(* IEC 61131-3 sources: volt/packages/volt-lsp-iec/test-corpus/pro2193/Device/Plc Logic/Application/09 Misc/Library Manager/CommFB, 61 files *)

(* ---- ADDR_TYPE.dut ---- *)
TYPE ADDR_TYPE :
UNION
	SYSTEM : IO_SYSTEM_TYPE;
	DP : DP_ADDR;
	PN : PN_ADDR;
END_UNION
END_TYPE

(* ---- AINFO_TYPE.dut ---- *)
TYPE AINFO_TYPE :
UNION
	DP : DP_AINFO;
	PN : PN_AINFO;
END_UNION
END_TYPE

(* ---- CNCT_STATE.dut ---- *)
TYPE CNCT_STATE :
(
	S1_INIT := 1,
	S2_IDLE := 2,
	S3_CONNECTING := 3,
	S4_CONNECTED := 4,
	S5_DISCONNECTING := 5,
	S6_ERROR := 6
);
END_TYPE

(* ---- DP_ADDR.dut ---- *)
TYPE DP_ADDR :
STRUCT
	SYSTEM : IO_SYSTEM_TYPE;
	VERSION : BYTE := 1;
	D : DP_DEVICE_ID;
	SLOT : BYTE;
END_STRUCT
END_TYPE

(* ---- DP_AINFO.dut ---- *)
TYPE DP_AINFO :
STRUCT
	D_LEN : BYTE;
	ATYPE : BYTE;
	SLOT : BYTE;
	ASPEC : BYTE;
	ADD_INFO : ARRAY [0..58] OF BYTE;
END_STRUCT
END_TYPE

(* ---- DP_DEVICE_ID.dut ---- *)
TYPE DP_DEVICE_ID :
STRUCT
	MASTER : BYTE;
	SEGMENT : BYTE;
	STATION : BYTE;
END_STRUCT
END_TYPE

(* ---- DP_DIAG.dut ---- *)
TYPE DP_DIAG :
STRUCT
	STATUS1 : IIoDrvProfibus.DP_StationStatus1;
	STATUS2 : IIoDrvProfibus.DP_StationStatus2;
	STATUS3 : IIoDrvProfibus.DP_StationStatus3;
	DIAG_MASTER_ADD : USINT;
	IDENT_NUMBER : UINT;
	EXTDIAG : ARRAY [0..235] OF BYTE;
END_STRUCT
END_TYPE

(* ---- ERRORCODE.dut ---- *)
TYPE ERRORCODE :
(
	NONE := 0,
	INVALID_ID := 16#40820000,
	UNKNOWN := 16#40000100,
	NOT_IMPLEMENTED := 16#40000101,
	RDIAG_PROFINET := 16#40000102,
	STACK_NOT_RUNNING := 16#40000103,
	NO_RESSOURCE := 16#40000104,
	BUFFER_SIZE := 16#40000105,
	INVALID_STATE := 16#40000110,
	ADDRESS_NOT_UNIQUE := 16#40000111,
	ADDRESS_INVALID := 16#40000112,
	DEVICE_NOT_FOUND := 16#40000113,
	DEVICETYPE_MISMATCH := 16#40000114,
	TIMEOUT := 16#40000115
);
END_TYPE

(* ---- ERRORCODE1_RW.dut ---- *)
TYPE ERRORCODE1_RW :
(
	INVALID_INDEX := 16#B0,
	WRITE_LENGTH_ERROR := 16#B1,
	INVALID_SLOT_OR_SUBSLOT := 16#B2,
	TYPE_CONFLICT := 16#B3,
	INVALID_AREA_OR_API := 16#B4,
	STATE_CONFLICT := 16#B5,
	ACCESS_DENIED := 16#B6,
	INVALID_RANGE := 16#B7,
	INVALID_PARAMETER := 16#B8,
	INVALID_TYPE := 16#B9,
	BACKUP := 16#BA
);
END_TYPE

(* ---- IO_SYSTEM_TYPE.dut ---- *)
TYPE IO_SYSTEM_TYPE :
(
	PROFIBUS_DP := 1,
	PROFINET_IO := 2
);
END_TYPE

(* ---- PN_ADDR.dut ---- *)
TYPE PN_ADDR :
STRUCT
	SYSTEM : IO_SYSTEM_TYPE;
	VERSION : BYTE := 1;
	MASTER : BYTE;
	D : PN_DEVICE_ID;
	API : DWORD;
	SLOT : WORD;
	SUBSLOT : WORD;
END_STRUCT
END_TYPE

(* ---- PN_AINFO.dut ---- *)
TYPE PN_AINFO :
STRUCT
	BLOCKTYPE : UINT;
	BLOCKLENGTH : UINT;
	VERSION : UINT;
	ALARMTYPE : UINT;
	API : UDINT;
	SLOT : UINT;
	SUBSLOT : UINT;
	MODULEIDENTNUMBER : UDINT;
	SUBMODULEIDENTNUMBER : UDINT;
	ALARMSPECIFIER : UINT;
	USI : UINT;
	ALARMDATA : ARRAY [0..(Constants.MAX_PN_ALARM_DATA - 1)] OF BYTE;
END_STRUCT
END_TYPE

(* ---- PN_DEVICE_ID.dut ---- *)
TYPE PN_DEVICE_ID :
STRUCT
	STATIONNAME : STRING;
	INSTANCE : WORD;
	DEVICE : WORD;
	VENDOR : WORD;
END_STRUCT
END_TYPE

(* ---- PRVREC_MODE.dut ---- *)
TYPE PRVREC_MODE :
(
	CHECK := 0,
	RECEIVE := 1,
	RECEIVE_BY_SLOT := 2,
	POS_RESPONSE := 3,
	NEG_RESPONSE := 4
);
END_TYPE

(* ---- PRVREC_STATE.dut ---- *)
TYPE PRVREC_STATE :
(
	S1_INIT,
	S2_IDLE,
	S3_ENABLED,
	S4_NEG_RESP,
	S5_RECEIVED,
	S6_CHECK,
	S7_POS_RESP,
	S8_NEG_RESP,
	S9_ERROR
);
END_TYPE

(* ---- RALARM_MODE.dut ---- *)
TYPE RALARM_MODE :
(
	ALL_ALARMS := 1,
	ALARM_BY_ID := 2,
	ALARM_BY_SLOT := 3,
	ALARM_BY_DEVICE := 4
);
END_TYPE

(* ---- RCVREC_MODE.dut ---- *)
TYPE RCVREC_MODE :
(
	CHECK := 0,
	RECEIVE := 1,
	RECEIVE_BY_SLOT := 2,
	POS_RESPONSE := 3,
	NEG_RESPONSE := 4
);
END_TYPE

(* ---- RCVREC_STATE.dut ---- *)
TYPE RCVREC_STATE :
(
	S1_INIT,
	S2_IDLE,
	S3_ENABLED,
	S4_NEG_RESP,
	S5_RECEIVED,
	S6_CHECK,
	S7_POS_RESP,
	S8_NEG_RESP,
	S9_ERROR
);
END_TYPE

(* ---- RDREC_STATE.dut ---- *)
TYPE RDREC_STATE :
(
	S1_INIT := 1,
	S2_IDLE := 2,
	S3_WAITING := 3,
	S4_HAVEDATA := 4,
	S5_ERROR := 5
);
END_TYPE

(* ---- READ_IND.dut ---- *)
TYPE READ_IND :
STRUCT
	SLOT : UINT;
	SUBSLOT : UINT;
	INDEX : UINT;
	RLEN : UINT;
	AR_ID : DWORD;
	SEQ_NUMBER : UINT;
END_STRUCT
END_TYPE

(* ---- SALRM_STATE.dut ---- *)
TYPE SALRM_STATE :
(
	S1_INIT,
	S2_IDLE,
	S3_WAITING,
	S4_HAVE_ACK,
	S5_ERROR
);
END_TYPE

(* ---- WRITE_IND.dut ---- *)
TYPE WRITE_IND :
STRUCT
	SLOT : UINT;
	SUBSLOT : UINT;
	INDEX : UINT;
	PRM : BOOL;
	AR_ID : DWORD;
	SEQ_NUMBER : UINT;
	LEN : UINT;
	DATA : POINTER TO BYTE;
END_STRUCT
END_TYPE

(* ---- WRREC_STATE.dut ---- *)
TYPE WRREC_STATE :
(
	S1_INIT := 1,
	S2_IDLE := 2,
	S3_WAITING := 3,
	S4_DATAWRITTEN := 4,
	S5_ERROR := 5
);
END_TYPE

(* ---- ADDRESSCONCEPT.gvl ---- *)
VAR_GLOBAL
	DUMMY : UDINT := 0;
END_VAR

(* ---- CONSTANTS.gvl ---- *)
VAR_GLOBAL
	INVALID_ID : UDINT := 16#FFFFFFFF;
	MAX_PN_ALARM_DATA : UDINT := 198;
END_VAR

(* ---- ICOMMFBALARMSENDER.itf ---- *)
INTERFACE ICOMMFBALARMSENDER
END_INTERFACE

METHOD ALARMCNF
VAR_INPUT
	ERROR : DWORD;
END_VAR
END_METHOD

(* ---- ICOMMFBCONNECTIONMANAGERFACTORY.itf ---- *)
INTERFACE ICOMMFBCONNECTIONMANAGERFACTORY
END_INTERFACE

METHOD GETCONNECTIONMANAGER : UDINT
VAR_INPUT
	CLIENT : IConnectionManagerClient;
END_VAR
VAR_OUTPUT
	CONNECTIONMANAGER : IConnectionManager;
END_VAR
VAR_IN_OUT
	D_ADDR : ADDR_TYPE;
END_VAR
END_METHOD

METHOD RELEASECONNECTIONMANAGER : UDINT
VAR_INPUT
	CLIENT : IConnectionManagerClient;
	CONNECTIONMANAGER : IConnectionManager;
END_VAR
END_METHOD

(* ---- ICOMMFBDIAGPROVIDER.itf ---- *)
INTERFACE ICOMMFBDIAGPROVIDER
END_INTERFACE

METHOD CHECKOWNER : BOOL
VAR_INPUT
	ID : UDINT;
END_VAR
END_METHOD

METHOD GETALARM : DWORD
VAR_INPUT
	MODE : INT;
	F_ID : DWORD;
END_VAR
VAR_OUTPUT
	NEW : BOOL;
	ID : DWORD;
	LEN : INT;
END_VAR
VAR_IN_OUT
	AINFO : AINFO_TYPE;
	CURRENTALARMID : UDINT;
END_VAR
END_METHOD

METHOD GETDIAG : DWORD
VAR_INPUT
	ID : DWORD;
END_VAR
VAR_OUTPUT
	BUSY : BOOL;
	LEN : INT;
END_VAR
VAR_IN_OUT
	DINFO : DP_DIAG;
END_VAR
END_METHOD

(* ---- ICOMMFBFACTORY.itf ---- *)
INTERFACE ICOMMFBFACTORY
END_INTERFACE

METHOD CHECKOWNER : BOOL
VAR_INPUT
	ID : UDINT;
END_VAR
END_METHOD

METHOD GETRDREC : POINTER TO RDRECBase
VAR_INPUT
	ID : UDINT;
END_VAR
VAR_IN_OUT
	CLIENT : RDREC;
END_VAR
END_METHOD

METHOD GETWRREC : POINTER TO WRRECBase
VAR_INPUT
	ID : UDINT;
END_VAR
VAR_IN_OUT
	CLIENT : WRREC;
END_VAR
END_METHOD

METHOD RELEASERDREC : BOOL
VAR_INPUT
	ID : UDINT;
END_VAR
VAR_IN_OUT
	CLIENT : RDREC;
END_VAR
END_METHOD

METHOD RELEASEWRREC : BOOL
VAR_INPUT
	ID : UDINT;
END_VAR
VAR_IN_OUT
	CLIENT : WRREC;
END_VAR
END_METHOD

(* ---- ICOMMFBFACTORYEXT.itf ---- *)
INTERFACE ICOMMFBFACTORYEXT
END_INTERFACE

METHOD TRYGETADDRESS : BOOL
VAR_INPUT
	ID : DWORD;
END_VAR
VAR_OUTPUT
	STATUS : DWORD;
END_VAR
VAR_IN_OUT
	ADDR : ADDR_TYPE;
END_VAR
END_METHOD

METHOD TRYGETID : BOOL
VAR_OUTPUT
	STATUS : DWORD;
	ID : DWORD;
END_VAR
VAR_IN_OUT
	ADDR : ADDR_TYPE;
END_VAR
END_METHOD

(* ---- ICOMMFBFACTORYIO.itf ---- *)
INTERFACE ICOMMFBFACTORYIO
END_INTERFACE

METHOD CHECKOWNER : BOOL
VAR_INPUT
	ID : UDINT;
END_VAR
END_METHOD

METHOD GETINPUTDATA : DWORD
VAR_INPUT
	ID : DWORD;
	OFFSET : UINT;
	LEN : UINT;
	INPUTS : POINTER TO BYTE;
END_VAR
VAR_OUTPUT
	IO_LEN : UINT;
	CONSISTENCY : BOOL;
END_VAR
END_METHOD

METHOD PUTOUTPUTDATA : DWORD
VAR_INPUT
	ID : DWORD;
	OFFSET : UINT;
	LEN : UINT;
	OUTPUTS : POINTER TO BYTE;
END_VAR
VAR_OUTPUT
	IO_LEN : UINT;
	CONSISTENCY : BOOL;
END_VAR
END_METHOD

(* ---- ICOMMFBFIELDDEVICE.itf ---- *)
INTERFACE ICOMMFBFIELDDEVICE
END_INTERFACE

METHOD ALARMREQ : DWORD
VAR_INPUT
	ALARMSENDER : ICommFBAlarmSender;
	ID : DWORD;
	ATYPE : UINT;
	ASPEC : UINT;
	LEN : UINT;
	AINFO : POINTER TO BYTE;
END_VAR
END_METHOD

METHOD CHECKREADIND : BOOL
VAR_INPUT
	MODE : UINT;
	F_ID : DWORD;
END_VAR
VAR_OUTPUT
	STATUS : DWORD;
	IND : Read_Ind;
END_VAR
END_METHOD

METHOD CHECKWRITEIND : BOOL
VAR_INPUT
	MODE : UINT;
	F_ID : DWORD;
END_VAR
VAR_OUTPUT
	STATUS : DWORD;
	IND : Write_Ind;
END_VAR
END_METHOD

METHOD READNEGRSP : DWORD
VAR_INPUT
	CODE1 : BYTE;
	CODE2 : BYTE;
END_VAR
VAR_IN_OUT
	IND : Read_Ind;
END_VAR
END_METHOD

METHOD READRSP : DWORD
VAR_INPUT
	LEN : UINT;
	RECORD : POINTER TO BYTE;
END_VAR
VAR_IN_OUT
	IND : Read_Ind;
END_VAR
END_METHOD

METHOD WRITENEGRSP : DWORD
VAR_INPUT
	CODE1 : BYTE;
	CODE2 : BYTE;
END_VAR
VAR_IN_OUT
	IND : Write_Ind;
END_VAR
END_METHOD

METHOD WRITERSP : DWORD
VAR_IN_OUT
	IND : Write_Ind;
END_VAR
END_METHOD

(* ---- ICONNECTIONMANAGER.itf ---- *)
INTERFACE ICONNECTIONMANAGER
END_INTERFACE

METHOD CONNECTREQ : DWORD
VAR_IN_OUT
	D_ADDR : ADDR_TYPE;
END_VAR
END_METHOD

METHOD RELEASEREQ : DWORD
END_METHOD

METHOD UPDATEADDRESS : DWORD
VAR_IN_OUT
	D_ADDR : ADDR_TYPE;
END_VAR
END_METHOD

(* ---- ICONNECTIONMANAGERCLIENT.itf ---- *)
INTERFACE ICONNECTIONMANAGERCLIENT
END_INTERFACE

METHOD CONNECTCNF
VAR_INPUT
	ID : DWORD;
	ERRORCODE : DWORD;
END_VAR
END_METHOD

METHOD ERRORIND
VAR_INPUT
	ERRORCODE : DWORD;
END_VAR
END_METHOD

METHOD RELEASECNF
VAR_INPUT
	ERRORCODE : DWORD;
END_VAR
END_METHOD

(* ---- IGENERICIDFACTORY.itf ---- *)
INTERFACE IGENERICIDFACTORY
END_INTERFACE

METHOD TRYGETIDFROMREFERENCE : BOOL
VAR_INPUT
	PREF : POINTER TO BYTE;
END_VAR
VAR_OUTPUT
	ID : DWORD;
END_VAR
END_METHOD

(* ---- ADDR.pou ---- *)
FUNCTION ADDR : DWORD
VAR_INPUT
	EN : BOOL := TRUE;
	ID : DWORD;
END_VAR
VAR_OUTPUT
	ENO : BOOL;
END_VAR
END_FUNCTION

(* ---- ID.pou ---- *)
FUNCTION ID : DWORD
VAR_INPUT
	EN : BOOL := TRUE;
	MASTER : BYTE;
	SEGMENT : BYTE;
	STATION : BYTE;
	SLOT : BYTE;
END_VAR
END_FUNCTION

(* ---- ID_FROM_REF.pou ---- *)
FUNCTION ID_FROM_REF : DWORD
VAR_INPUT
	PREF : POINTER TO BYTE;
END_VAR
END_FUNCTION

(* ---- SLOT_ID.pou ---- *)
FUNCTION SLOT_ID : DWORD
VAR_INPUT
	EN : BOOL := TRUE;
	ID : DWORD;
	SLOT : BYTE;
END_VAR
VAR_OUTPUT
	ENO : BOOL;
END_VAR
END_FUNCTION

(* ---- SUBSLOT_ID.pou ---- *)
FUNCTION SUBSLOT_ID : DWORD
VAR_INPUT
	EN : BOOL := TRUE;
	ID : DWORD;
	SLOT : UINT;
	SUBSLOT : UINT;
END_VAR
VAR_OUTPUT
	ENO : BOOL;
END_VAR
END_FUNCTION

(* ---- ADDR_TO_ID.pou ---- *)
FUNCTION_BLOCK ADDR_TO_ID
VAR_INPUT
	EN : BOOL := TRUE;
END_VAR
VAR_OUTPUT
	ENO : BOOL;
	STATUS : DWORD;
	ID : DWORD;
END_VAR
VAR_IN_OUT
	ADDR : ADDR_TYPE;
END_VAR
VAR
	S_INSTANCEHANDLER : InstanceHandler;
	I : DINT;
END_VAR
END_FUNCTION_BLOCK

(* ---- ALARMSENDERINTERNAL.pou ---- *)
FUNCTION_BLOCK ALARMSENDERINTERNAL
VAR_INPUT
	SALARM : POINTER TO SALARM;
END_VAR
END_FUNCTION_BLOCK

METHOD ALARMCNF
VAR_INPUT
	ERROR : DWORD;
END_VAR
END_METHOD

(* ---- CNCT.pou ---- *)
FUNCTION_BLOCK CNCT
VAR_INPUT
	REQ : BOOL;
	D_ADDR : ADDR_TYPE;
END_VAR
VAR_OUTPUT
	VALID : BOOL;
	ERROR : BOOL;
	BUSY : BOOL;
	STATUS : DWORD;
	ID : DWORD := Constants.INVALID_ID;
END_VAR
VAR
	S_INSTANCEHANDLER : InstanceHandler;
	_FACTORY : ICommFBConnectionManagerFactory;
	_CONNECTIONMANAGER : IConnectionManager;
	_REQ : BOOL;
	_STATE : CNCT_State := CNCT_State.S2_Idle;
	_ERRORCODE : UDINT;
	_CONNECTREQ : UDINT;
	_CONNECTID : DWORD := Constants.INVALID_ID;
	_RECVCONNECTCNF : BOOL;
	_RECVRELEASECNF : BOOL;
	_RECVABORTIND : BOOL;
	_CLIENT : ConnectionManagerClientInternal;
END_VAR
END_FUNCTION_BLOCK

METHOD ABORTIND
VAR_INPUT
	ERRORCODE : DWORD;
END_VAR
END_METHOD

METHOD CONNECTCNF
VAR_INPUT
	ID : DWORD;
	ERRORCODE : DWORD;
END_VAR
END_METHOD

METHOD RELEASECNF
VAR_INPUT
	ERRORCODE : DWORD;
END_VAR
END_METHOD

(* ---- CONNECTIONMANAGERCLIENTIMPLICITID.pou ---- *)
FUNCTION_BLOCK CONNECTIONMANAGERCLIENTIMPLICITID
VAR_INPUT
	CNCT : POINTER TO CREATE_ID;
END_VAR
END_FUNCTION_BLOCK

METHOD CONNECTCNF
VAR_INPUT
	ID : DWORD;
	ERRORCODE : DWORD;
END_VAR
END_METHOD

METHOD ERRORIND
VAR_INPUT
	ERRORCODE : DWORD;
END_VAR
END_METHOD

METHOD RELEASECNF
VAR_INPUT
	ERRORCODE : DWORD;
END_VAR
END_METHOD

(* ---- CONNECTIONMANAGERCLIENTINTERNAL.pou ---- *)
FUNCTION_BLOCK CONNECTIONMANAGERCLIENTINTERNAL
VAR_INPUT
	CNCT : POINTER TO CNCT;
END_VAR
END_FUNCTION_BLOCK

METHOD CONNECTCNF
VAR_INPUT
	ID : DWORD;
	ERRORCODE : DWORD;
END_VAR
END_METHOD

METHOD ERRORIND
VAR_INPUT
	ERRORCODE : DWORD;
END_VAR
END_METHOD

METHOD RELEASECNF
VAR_INPUT
	ERRORCODE : DWORD;
END_VAR
END_METHOD

(* ---- CREATE_ID.pou ---- *)
FUNCTION_BLOCK CREATE_ID
VAR_INPUT
	EN : BOOL := TRUE;
END_VAR
VAR_OUTPUT
	ENO : BOOL;
	STATUS : DWORD;
	ID : DWORD;
END_VAR
VAR_IN_OUT
	ADDR : ADDR_TYPE;
END_VAR
VAR
	S_INSTANCEHANDLER : InstanceHandler;
	_FACTORY : ICommFBConnectionManagerFactory;
	_CONNECTIONMANAGER : IConnectionManager;
	_STATE : CNCT_State := CNCT_State.S2_Idle;
	_ERRORCODE : UDINT;
	_CONNECTID : DWORD := Constants.INVALID_ID;
	_RECVCONNECTCNF : BOOL;
	_RECVRELEASECNF : BOOL;
	_RECVABORTIND : BOOL;
	_CLIENT : ConnectionManagerClientImplicitID;
	D_ADDR : ADDR_TYPE;
END_VAR
END_FUNCTION_BLOCK

METHOD ABORTIND
VAR_INPUT
	ERRORCODE : DWORD;
END_VAR
END_METHOD

METHOD CONNECTCNF
VAR_INPUT
	ID : DWORD;
	ERRORCODE : DWORD;
END_VAR
END_METHOD

METHOD RELEASECNF
VAR_INPUT
	ERRORCODE : DWORD;
END_VAR
END_METHOD

(* ---- GETIO_PART.pou ---- *)
FUNCTION_BLOCK GETIO_PART
VAR_INPUT
	EN : BOOL;
	ID : DWORD;
	OFFSET : INT;
	LEN : INT;
	INPUTS : POINTER TO BYTE;
END_VAR
VAR_OUTPUT
	ENO : BOOL;
	STATUS : DWORD;
	ERROR : BOOL;
END_VAR
VAR
	S_INSTANCEHANDLER : InstanceHandler;
	I : DINT;
	_FACTORY : ICommFBFactoryIO;
	IOLEN : UINT;
	TRANSFERCONSISTENT : BOOL;
END_VAR
END_FUNCTION_BLOCK

(* ---- ID_TO_ADDR.pou ---- *)
FUNCTION_BLOCK ID_TO_ADDR
VAR_INPUT
	EN : BOOL := TRUE;
	ID : DWORD;
END_VAR
VAR_OUTPUT
	ENO : BOOL;
	STATUS : DWORD;
END_VAR
VAR_IN_OUT
	ADDR : ADDR_TYPE;
END_VAR
VAR
	S_INSTANCEHANDLER : InstanceHandler;
	I : DINT;
	FACTORY : ICommFBFactoryExt;
END_VAR
END_FUNCTION_BLOCK

(* ---- INSTANCEHANDLER.pou ---- *)
FUNCTION_BLOCK INSTANCEHANDLER
VAR
	S_INSTANCECOUNT : UINT;
	S_FACTORIES : ARRAY [0..(MAX_INSTANCES - 1)] OF ICommFBFactory;
	S_FACTORIESEXT : ARRAY [0..(MAX_INSTANCES - 1)] OF ICommFBFactoryExt;
	S_FACTORIESIO : ARRAY [0..(MAX_INSTANCES - 1)] OF ICommFBFactoryIO;
	S_FACTORIESCONNECTIONS : ARRAY [0..(MAX_INSTANCES - 1)] OF ICommFBConnectionManagerFactory;
	S_FIELDDEVICES : ARRAY [0..(MAX_INSTANCES - 1)] OF ICommFBFieldDevice;
	S_GENERICIDFACTORIES : ARRAY [0..(MAX_INSTANCES - 1)] OF IGenericIDFactory;
	S_IDS : UDINT := (MAX_INSTANCES - 1);
	S_DIAGPROVIDERS : ARRAY [0..(MAX_INSTANCES - 1)] OF ICommFBDiagProvider;
	MAX_INSTANCES : UINT := 8;
END_VAR
END_FUNCTION_BLOCK

METHOD CREATEID : UDINT
END_METHOD

METHOD GETCONNECTIONMANAGERFACTORY : UDINT
VAR_OUTPUT
	FACTORY : ICommFBConnectionManagerFactory;
END_VAR
VAR_IN_OUT
	D_ADDR : ADDR_TYPE;
END_VAR
END_METHOD

METHOD GETDIAGFACTORY : UDINT
VAR_INPUT
	ID : UDINT;
END_VAR
VAR_OUTPUT
	DIAGPROVIDER : ICommFBDiagProvider;
END_VAR
END_METHOD

METHOD GETFACTORY : ICommFBFactory
VAR_INPUT
	ID : UDINT;
END_VAR
END_METHOD

METHOD GETFIELDDEVICE : DWORD
VAR_INPUT
	ID : UDINT;
END_VAR
VAR_OUTPUT
	FIELDDEVICE : ICommFBFieldDevice;
END_VAR
END_METHOD

METHOD GETIOFACTORY : UDINT
VAR_INPUT
	ID : UDINT;
END_VAR
VAR_OUTPUT
	FACTORY : ICommFBFactoryIO;
END_VAR
END_METHOD

METHOD REGISTER : UINT
VAR_INPUT
	FACTORY : ICommFBFactory;
END_VAR
END_METHOD

METHOD REGISTERDIAG : UINT
VAR_INPUT
	FACTORY : ICommFBFactory;
	DIAGPROVIDER : ICommFBDiagProvider;
END_VAR
END_METHOD

METHOD REGISTEREXT : UINT
VAR_INPUT
	FACTORY : ICommFBFactory;
	DIAGPROVIDER : ICommFBDiagProvider;
	FACTORYEXT : ICommFBFactoryExt;
END_VAR
END_METHOD

METHOD REGISTEREXTIO : UINT
VAR_INPUT
	FACTORY : ICommFBFactory;
	DIAGPROVIDER : ICommFBDiagProvider;
	FACTORYEXT : ICommFBFactoryExt;
	UPDATEIO : ICommFBFactoryIO;
END_VAR
END_METHOD

METHOD REGISTERFIELDDEVICE : UINT
VAR_INPUT
	FACTORY : ICommFBFactory;
	FACTORYEXT : ICommFBFactoryExt;
	DEVICE : ICommFBFieldDevice;
END_VAR
END_METHOD

METHOD REGISTERINTERFACES : UINT
VAR_INPUT
	FACTORY : ICommFBFactory;
	DIAGPROVIDER : ICommFBDiagProvider;
	FACTORYEXT : ICommFBFactoryExt;
	UPDATEIO : ICommFBFactoryIO;
	CNCT : ICommFBConnectionManagerFactory;
END_VAR
END_METHOD

(* ---- PRVREC.pou ---- *)
FUNCTION_BLOCK PRVREC
VAR_INPUT
	EN : BOOL;
	MODE : UINT;
	F_ID : DWORD;
	CODE1 : BYTE;
	CODE2 : BYTE;
	LEN : UINT;
	RECORD : POINTER TO BYTE;
END_VAR
VAR_OUTPUT
	ENO : BOOL;
	NEW : BOOL;
	STATUS : DWORD;
	SLOT : UINT;
	SUBSLOT : UINT;
	INDEX : UINT;
	RLEN : UINT;
END_VAR
VAR
	S_INSTANCEHANDLER : InstanceHandler;
	_STATE : PRVREC_State := PRVREC_State.S1_INIT;
	_DEVICE : ICommFBFieldDevice;
	_READIND : Read_Ind;
	EMPTYIND : Read_Ind;
END_VAR
END_FUNCTION_BLOCK

(* ---- RALARM.pou ---- *)
FUNCTION_BLOCK RALARM
VAR_INPUT
	EN : BOOL;
	MODE : INT;
	F_ID : DWORD;
END_VAR
VAR_OUTPUT
	ENO : BOOL;
	NEW : BOOL;
	STATUS : DWORD;
	ID : DWORD;
	LEN : INT;
END_VAR
VAR_IN_OUT
	AINFO : AINFO_TYPE;
END_VAR
VAR
	S_INSTANCEHANDLER : InstanceHandler;
	M_EN : BOOL;
	M_MODE : INT;
	M_F_ID : DWORD;
	M_FACTORY : ICommFBDiagProvider;
	M_CURRENTALARMID : UDINT := Constants.INVALID_ID;
END_VAR
END_FUNCTION_BLOCK

(* ---- RCVREC.pou ---- *)
FUNCTION_BLOCK RCVREC
VAR_INPUT
	EN : BOOL;
	MODE : UINT;
	F_ID : DWORD;
	MLEN : UINT;
	CODE1 : BYTE;
	CODE2 : BYTE;
	RECORD : POINTER TO BYTE;
END_VAR
VAR_OUTPUT
	ENO : BOOL;
	NEW : BOOL;
	STATUS : DWORD;
	SLOT : UINT;
	SUBSLOT : UINT;
	INDEX : UINT;
	LEN : UINT;
END_VAR
VAR
	S_INSTANCEHANDLER : InstanceHandler;
	_STATE : RCVREC_State := RCVREC_State.S1_INIT;
	_DEVICE : ICommFBFieldDevice;
	_WRITEIND : Write_Ind;
	EMPTYIND : Write_Ind;
	I : DINT;
END_VAR
END_FUNCTION_BLOCK

(* ---- RDIAG.pou ---- *)
FUNCTION_BLOCK RDIAG
VAR_INPUT
	REQ : BOOL;
	ID : DWORD;
	MLEN : INT;
END_VAR
VAR_OUTPUT
	VALID : BOOL;
	BUSY : BOOL;
	ERROR : BOOL;
	STATUS : DWORD;
	LEN : INT;
END_VAR
VAR_IN_OUT
	DINFO : DP_DIAG;
END_VAR
VAR
	S_INSTANCEHANDLER : InstanceHandler;
	M_FACTORY : ICommFBDiagProvider;
END_VAR
END_FUNCTION_BLOCK

(* ---- RDREC.pou ---- *)
FUNCTION_BLOCK RDREC
VAR_INPUT
	REQ : BOOL;
	ID : DWORD;
	INDEX : INT;
	MLEN : INT;
	RECORD : POINTER TO BYTE;
END_VAR
VAR_OUTPUT
	VALID : BOOL;
	BUSY : BOOL;
	ERROR : BOOL;
	STATUS : DWORD;
	LEN : INT;
END_VAR
VAR
	M_FACTORY : ICommFBFactory;
	M_PRDREC : POINTER TO RDRECbase;
	_REQ : BOOL;
	S_INSTANCEHANDLER : InstanceHandler;
END_VAR
END_FUNCTION_BLOCK

(* ---- RDRECBASE.pou ---- *)
FUNCTION_BLOCK RDRECBASE
VAR_INPUT
	REQ : BOOL;
	ID : DWORD;
	INDEX : INT;
	MLEN : INT;
	RECORD : POINTER TO BYTE;
END_VAR
VAR_OUTPUT
	VALID : BOOL;
	ERROR : BOOL;
	BUSY : BOOL;
	STATUS : DWORD;
	LEN : INT;
END_VAR
END_FUNCTION_BLOCK

(* ---- RDRECDEFAULT.pou ---- *)
FUNCTION_BLOCK RDRECDEFAULT EXTENDS RDRECbase
VAR
	STATE : RDREC_State := RDREC_State.S2_Idle;
	_ERRORCODE : UDINT;
	DATALEN : INT;
	PRECORDDATA : POINTER TO BYTE;
	NEXT : BOOL;
END_VAR
END_FUNCTION_BLOCK

METHOD COPYDATA
VAR_INPUT
	LENGTH : INT;
	PDATA : POINTER TO BYTE;
END_VAR
END_METHOD

METHOD NEGRESPONSE
VAR_INPUT
	ERRORCODE : DWORD;
END_VAR
END_METHOD

METHOD POSRESPONSE
END_METHOD

METHOD START : UDINT
END_METHOD

METHOD WAITING
END_METHOD

(* ---- SALARM.pou ---- *)
FUNCTION_BLOCK SALARM
VAR_INPUT
	REQ : BOOL;
	ID : DWORD;
	ATYPE : UINT;
	ASPEC : UINT;
	LEN : UINT;
	AINFO : POINTER TO BYTE;
END_VAR
VAR_OUTPUT
	DONE : BOOL;
	BUSY : BOOL;
	ERROR : BOOL;
	STATUS : DWORD;
END_VAR
VAR
	S_INSTANCEHANDLER : InstanceHandler;
	_REQ : BOOL;
	_STATE : SALRM_State := SALRM_State.S1_INIT;
	SEND_RESULT : UDINT;
	_DEVICE : ICommFBFieldDevice;
	_CLIENT : AlarmSenderInternal;
	_ERROR : DWORD;
	_CONTINUE : BOOL;
END_VAR
END_FUNCTION_BLOCK

METHOD ALARMCNF
VAR_INPUT
	ERROR : DWORD;
END_VAR
END_METHOD

METHOD NEG_RESPONSE
VAR_INPUT
	ERROR : DWORD;
END_VAR
END_METHOD

METHOD POS_RESPONSE
END_METHOD

(* ---- SETIO_PART.pou ---- *)
FUNCTION_BLOCK SETIO_PART
VAR_INPUT
	EN : BOOL;
	ID : DWORD;
	OFFSET : INT;
	LEN : INT;
	OUTPUTS : POINTER TO BYTE;
END_VAR
VAR_OUTPUT
	ENO : BOOL;
	STATUS : DWORD;
	ERROR : BOOL;
END_VAR
VAR
	S_INSTANCEHANDLER : InstanceHandler;
	I : DINT;
	_FACTORY : ICommFBFactoryIO;
	IOLEN : UINT;
	TRANSFERCONSISTENT : BOOL;
END_VAR
END_FUNCTION_BLOCK

(* ---- WRREC.pou ---- *)
FUNCTION_BLOCK WRREC
VAR_INPUT
	REQ : BOOL;
	ID : DWORD;
	INDEX : INT;
	LEN : INT;
	RECORD : POINTER TO BYTE;
END_VAR
VAR_OUTPUT
	DONE : BOOL;
	BUSY : BOOL;
	ERROR : BOOL;
	STATUS : DWORD;
END_VAR
VAR
	M_FACTORY : ICommFBFactory;
	M_PWRREC : POINTER TO WRRECbase;
	_REQ : BOOL;
	S_INSTANCEHANDLER : InstanceHandler;
END_VAR
END_FUNCTION_BLOCK

(* ---- WRRECBASE.pou ---- *)
FUNCTION_BLOCK WRRECBASE
VAR_INPUT
	REQ : BOOL;
	ID : DWORD;
	INDEX : INT;
	LEN : INT;
	RECORD : POINTER TO BYTE;
END_VAR
VAR_OUTPUT
	DONE : BOOL;
	BUSY : BOOL;
	ERROR : BOOL;
	STATUS : DWORD;
END_VAR
END_FUNCTION_BLOCK

(* ---- WRRECDEFAULT.pou ---- *)
FUNCTION_BLOCK WRRECDEFAULT EXTENDS WRRECbase
VAR
	STATE : WRREC_State := WRREC_State.S2_Idle;
	ERRORCODE : UDINT;
END_VAR
END_FUNCTION_BLOCK

METHOD NEGRESPONSE
VAR_INPUT
	ERRORCODE : DWORD;
END_VAR
END_METHOD

METHOD POSRESPONSE
END_METHOD

METHOD START : UDINT
END_METHOD

METHOD WAITING
END_METHOD
